(* IEC 61131-3 sources: kns-pump-station/tests/POUs/Model/FB_ScaledClock_Test, 10 files *)

(* ---- FB_ScaledClock_Test.decl.st ---- *)
// Назначение: набор coUnit для FB_ScaledClock — часы контура с ускорением: совпадение с системным
//             временем при k = 1, ограничение и неконечный коэффициент, монотонность при смене k, отношение
//             интервалов k (оценка «вилкой» по системному времени, без ожидания), ручной режим.
//             Реальное время читается только в проверках, которые ничего не ждут (docs/TESTING.md библиотеки).
// Автор:      kr0nsch
// Версия:     0.1.0
// Документ:   docs/DESIGN.md, разделы 11.3, 14.1
FUNCTION_BLOCK FB_ScaledClock_Test EXTENDS coUnit.FB_TestSuite
VAR CONSTANT
    R_SCALE_MAX : REAL := 50.0;           // SIM_TIME_SCALE_MAX
    LR_ROUND_NS : LREAL := 2.0;           // округление LREAL → LTIME двух отметок, нс
    LT_MANUAL_START : LTIME := LTIME#2H;
    LT_MANUAL_STEP : LTIME := LTIME#1S500MS;
    LT_MANUAL_AFTER : LTIME := LTIME#2H1S500MS;
    UI_READS : UINT := 1000;              // чтений часов в проверке монотонности
    DW_NAN : DWORD := 16#7FC00000;        // тихий NaN
    DW_INF : DWORD := 16#7F800000;        // +∞
    DW_NEG_INF : DWORD := 16#FF800000;    // −∞
END_VAR

(* ---- AdvanceIgnoredOutsideManual.method.decl.st ---- *)
// AdvanceL вне ручного режима ничего не делает: часы по-прежнему равны системному времени (k = 1).
METHOD PRIVATE AdvanceIgnoredOutsideManual
VAR
    fbClock : FB_ScaledClock;
    ltR0 : LTIME;
    ltR1 : LTIME;
    ltNow : LTIME;
END_VAR

(* ---- DefaultsScaleOneAndSystemTime.method.decl.st ---- *)
// Без Update: коэффициент 1, Now() — системное время (между двумя чтениями LTIME()).
METHOD PRIVATE DefaultsScaleOneAndSystemTime
VAR
    fbClock : FB_ScaledClock;   // проверяемые часы
    ltR0 : LTIME;               // системное время до чтения часов
    ltR1 : LTIME;               // после
    ltNow : LTIME;              // показание часов
END_VAR

(* ---- ManualAdvance.method.decl.st ---- *)
// Ручной режим: Now() = заданное время, меняется только AdvanceL, коэффициент не влияет; после
// выключения часы продолжают от ручного времени (не назад).
METHOD PRIVATE ManualAdvance
VAR
    fbClock : FB_ScaledClock;
    ltR0 : LTIME;
    ltR1 : LTIME;
    ltNow : LTIME;
END_VAR

(* ---- NanScaleIsOne.method.decl.st ---- *)
// Неконечный коэффициент (NaN, ±∞) — 1.
METHOD PRIVATE NanScaleIsOne
VAR
    fbClock : FB_ScaledClock;
    uBits : PL.U_RealBits;      // неконечные значения REAL по битам
END_VAR

(* ---- ScaleChangeIsMonotonic.method.decl.st ---- *)
// Смена коэффициента 1 → 50 → 1 → 20 перебазирует часы: время не идёт назад.
METHOD PRIVATE ScaleChangeIsMonotonic
VAR
    fbClock : FB_ScaledClock;
    altRead : ARRAY[1..6] OF LTIME;     // показания после каждой смены
END_VAR

(* ---- ScaleClampedToMax.method.decl.st ---- *)
// Коэффициент ограничивается 1…SIM_TIME_SCALE_MAX.
METHOD PRIVATE ScaleClampedToMax
VAR
    fbClock : FB_ScaledClock;
END_VAR

(* ---- ScaleFiftyBracketsRealTime.method.decl.st ---- *)
// k = 50: интервал часов между двумя чтениями лежит в «вилке» 50 · (интервал системного времени),
// посчитанной по чтениям LTIME() до и после каждого показания; часы монотонны (1000 чтений подряд).
METHOD PRIVATE ScaleFiftyBracketsRealTime
VAR
    fbClock : FB_ScaledClock;
    ltRa0 : LTIME;              // системное время вокруг первого показания
    ltRa1 : LTIME;
    ltRb0 : LTIME;              // вокруг второго
    ltRb1 : LTIME;
    ltSa : LTIME;               // показания часов
    ltSb : LTIME;
    ltPrev : LTIME;
    ltCur : LTIME;
    uiI : UINT;
    xMono : BOOL := TRUE;       // все чтения не убывают
    lrScaled_ns : LREAL;        // интервал часов
    lrLow_ns : LREAL;           // нижняя граница вилки
    lrHigh_ns : LREAL;          // верхняя граница
END_VAR

(* ---- ScaleFiftyBracketsRealTime.method.impl.st ---- *)
coUnit.TEST('ScaledClock_ScaleFiftyBracketsRealTime');

fbClock.Update(rTimeScale := R_SCALE_MAX);
ltRa0 := LTIME();
ltSa := fbClock.Now();
ltRa1 := LTIME();
ltPrev := ltSa;
FOR uiI := 1 TO UI_READS DO
    ltCur := fbClock.Now();
    xMono := xMono AND ltCur >= ltPrev;
    ltPrev := ltCur;
END_FOR
ltRb0 := LTIME();
ltSb := fbClock.Now();
ltRb1 := LTIME();
AssertTrue(Condition := xMono AND ltSb >= ltSa, Message := 'k = 50: clock is monotonic');
lrScaled_ns := ULINT_TO_LREAL(LTIME_TO_ULINT(ltSb - ltSa));
lrLow_ns := REAL_TO_LREAL(R_SCALE_MAX) * ULINT_TO_LREAL(LTIME_TO_ULINT(ltRb0 - ltRa1));
lrHigh_ns := REAL_TO_LREAL(R_SCALE_MAX) * ULINT_TO_LREAL(LTIME_TO_ULINT(ltRb1 - ltRa0));
AssertTrue(Condition := lrScaled_ns >= lrLow_ns - LR_ROUND_NS AND lrScaled_ns <= lrHigh_ns + LR_ROUND_NS,
           Message := 'k = 50: clock interval is 50 x system interval');

coUnit.TEST_FINISHED();

(* ---- ScaleOneEqualsSystem.method.decl.st ---- *)
// k = 1: часы совпадают с LTIME() и после нескольких чтений.
METHOD PRIVATE ScaleOneEqualsSystem
VAR
    fbClock : FB_ScaledClock;
    ltR0 : LTIME;
    ltR1 : LTIME;
    ltNow : LTIME;
END_VAR
